DATA_BLOCK "GDB_FraktalHal"
{ S7_Optimized_Access := 'TRUE' }
VERSION : 0.1
NON_RETAIN
VAR
    Data {ExternalAccessible := 'False'; ExternalVisible := 'False'; ExternalWritable := 'False'} : "ST_FraktalHal";
END_VAR
BEGIN
END_DATA_BLOCK
